// TIA Portal V15.1 export
// export: Created 2026-11-02T18:55:12.3174301Z, ExportSetting WithDefaults, DisplayName Totally Integrated Automation Portal, DisplayVersion V15.1, DisplayName TIA Portal Openness, DisplayVersion V15.1, DisplayName STEP 7 Professional, DisplayVersion V15.1, DisplayName WinCC Professional, DisplayVersion V15.1
VAR_GLOBAL   // PLC tag table "Tag table_1"
END_VAR
